Fanuc KAREL source: ke00001.KL

-- PROVISIONAL review KL for V1013-1; original PC SHA256 72bdec58595e4dd009d3b9b828a888123a85489eed0b3d0a45762380532b6f22
-- Incomplete behavior may be omitted. Consult companion uncertainty JSON. Do not deploy.
PROGRAM KE00001
%NOLOCKGROUP
BEGIN
  -- UNRESOLVED_PC offsets 5-12; opcodes 9D,23
  -- UNRESOLVED_PC offsets 17-41; opcodes 27,22,22,2A,22,31
  -- UNRESOLVED_PC offsets 46-50; opcodes 7F
END KE00001
